{attribute 'qualified_only'}
{attribute 'strict'}
TYPE E_TankFault :
(
    None           := 0,
    EStop          := 1,
    BusFault       := 2,
    SensorMismatch := 3,
    FillTimeout    := 4,
    DrainTimeout   := 5
) INT;
END_TYPE

(* stored: Version 1.1.0.1
   DUT E_TankFault: Id {3531d4e4-ab6b-428f-873d-adf9bcb118a3} *)
